(* IEC 61131-3 sources: nautilus/siemens/writer/testdata/arrays, 2 files *)

(* ---- lib.st ---- *)
TYPE
  R : STRUCT
    n : STRING;
    v : REAL := 1.5;
    hist : ARRAY[0..2] OF INT;
  END_STRUCT;
  Mode : (Idle, Run := 5) := Run;
END_TYPE

VAR_GLOBAL CONSTANT
  STAGES : INT := 2 + 1;
END_VAR

FUNCTION Pick : REAL
VAR_INPUT k : INT; t : ARRAY[1..3] OF REAL; END_VAR
Pick := t[k];
END_FUNCTION

FUNCTION_BLOCK Grid
VAR_INPUT k : INT; x : REAL; END_VAR
VAR_OUTPUT y : REAL; END_VAR
VAR tbl : ARRAY[-2..2, 0..3] OF REAL; END_VAR
tbl[k, k + 1] := x;
y := tbl[k, k + 1];
END_FUNCTION_BLOCK

FUNCTION_BLOCK Outer
VAR_INPUT k : INT; END_VAR
VAR_OUTPUT y : REAL; END_VAR
VAR g : Grid; END_VAR
g(k := k, x := 2.0, y => y);
END_FUNCTION_BLOCK

(* ---- Main.st ---- *)
PROGRAM Main
VAR CONSTANT N : INT := 4; END_VAR
VAR_EXTERNAL sel : INT; tbl : ARRAY[1..3] OF REAL; END_VAR
VAR
  a : ARRAY[1..N] OF DINT;
  b : ARRAY[-2..2, 0..3] OF INT;
  r : ARRAY[1..STAGES] OF R;
  m : ARRAY[0..1] OF Mode;
  s : ARRAY[1..2] OF STRING;
  i, j : INT;
  sum : DINT;
  x, y : REAL;
  act : R;
  inst : Grid;
  o : Outer;
  outs : ARRAY[0..2] OF REAL;
END_VAR
FOR i := 1 TO N DO a[i] := i; sum := sum + a[i]; END_FOR;
a[2] := 7;
b[i, j + 1] := b[-2, 0];
act := r[sel];
r[1].hist[j] := i;
x := tbl[i] + Pick(k := j, t := tbl) * 2.0;
inst(k := sel, x := tbl[j], y => outs[i]);
o(k := j, y => y);
IF x > 0.0 THEN y := 1.0; ELSIF tbl[j] > 1.0 THEN y := 2.0; ELSE y := 3.0; END_IF;
WHILE a[i] > 0 DO i := i + 1; END_WHILE;
outs[i] := tbl[j] + Pick(k := i, t := tbl);
s[1] := 'x';
m[0] := Idle;
END_PROGRAM
